// TIA Portal V17 export
// export: Created 2026-11-08T05:50:28.1424478Z, ExportSetting WithDefaults, DisplayName Totally Integrated Automation Portal, DisplayVersion V17, DisplayName TIA Portal Openness, DisplayVersion V17, DisplayName TIA Portal Version Control Interface, DisplayVersion V17, DisplayName STEP 7 Professional, DisplayVersion V17, DisplayName STEP 7 Safety, DisplayVersion V17, DisplayName WinCC Professional, DisplayVersion V17
DATA_BLOCK "DB_Motor_Mealy"   // DB5
VERSION : 0.1
// stored: AutoNumber true, DBAccessibleFromOPCUA true, InstanceOfName FB_Motor_Mealy, InstanceOfType FB
"FB_Motor_Mealy"
   // VAR_INPUT
   //    Marcha : Bool;
   //    Paro : Bool;
   //    Termico_OK : Bool;
   //    Reset : Bool;
   // END_VAR
   // VAR_OUTPUT
   //    Motor : Bool;
   //    Piloto_Marcha : Bool;
   //    Piloto_Falla : Bool;
   //    Estado : Int;
   // END_VAR
   // VAR
   //    Estado_Actual : Int;
   // END_VAR
BEGIN
END_DATA_BLOCK
